Staubli VAL3: getSize.pgx

public program getSize(num& x_nSize)
begin
  // give back the size to trajectory field
  x_nSize=size(trajTemp:tTrajItem)
end
